FUNCTION_BLOCK FB_Startup
VAR_INPUT
END_VAR
VAR_OUTPUT
END_VAR
VAR
	timer1 : TON;
	timer2 : TON;
	timer3 : TON;
	timer4 : TON;
	timer5 : TON;
	timer6 : TON;
	timer7 : TON;
	EMG_STOP_RELEASED : BOOL;
END_VAR

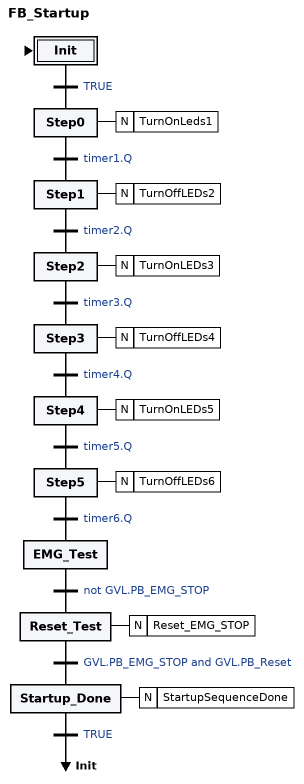
INITIAL_STEP Init:
END_STEP
TRANSITION FROM Init TO Step0
    := TRUE;
END_TRANSITION
STEP Step0:
    TurnOnLeds1(N);
END_STEP
TRANSITION FROM Step0 TO Step1
    := timer1.Q;
END_TRANSITION
STEP Step1:
    TurnOffLEDs2(N);
END_STEP
TRANSITION FROM Step1 TO Step2
    := timer2.Q;
END_TRANSITION
STEP Step2:
    TurnOnLEDs3(N);
END_STEP
TRANSITION FROM Step2 TO Step3
    := timer3.Q;
END_TRANSITION
STEP Step3:
    TurnOffLEDs4(N);
END_STEP
TRANSITION FROM Step3 TO Step4
    := timer4.Q;
END_TRANSITION
STEP Step4:
    TurnOnLEDs5(N);
END_STEP
TRANSITION FROM Step4 TO Step5
    := timer5.Q;
END_TRANSITION
STEP Step5:
    TurnOffLEDs6(N);
END_STEP
TRANSITION FROM Step5 TO EMG_Test
    := timer6.Q;
END_TRANSITION
STEP EMG_Test:
END_STEP
TRANSITION FROM EMG_Test TO Reset_Test
    := not GVL.PB_EMG_STOP;
END_TRANSITION
STEP Reset_Test:
    Reset_EMG_STOP(N);
END_STEP
TRANSITION FROM Reset_Test TO Startup_Done
    := GVL.PB_EMG_STOP and GVL.PB_Reset;
END_TRANSITION
STEP Startup_Done:
    StartupSequenceDone(N);
END_STEP
TRANSITION FROM Startup_Done TO Init
    := TRUE;
END_TRANSITION

METHOD AllLEDsTrigger : BOOL
VAR_INPUT
	OnOff : BOOL; // OnOff - Turn off, True - Turn On
END_VAR
GVL.LED_Comm_Fault := OnOff;
GVL.LED_EE_Grip := OnOff;
GVL.LED_EE_Ungrip := OnOff;
GVL.LED_EMG_STOP := OnOff;
GVL.LED_J1_CCW := OnOff;
GVL.LED_J1_CW := OnOff;
GVL.LED_J2_CCW := OnOff;
GVL.LED_J2_CW := OnOff;
GVL.LED_J3_CCW := OnOff;
GVL.LED_J3_CW := OnOff;
GVL.LED_Record_Delay := OnOff;
GVL.LED_Record_Pos := OnOff;
GVL.LED_Reset := OnOff;
GVL.LED_Start_Pause := OnOff;
GVL.LED_Warning := OnOff;
END_METHOD

ACTION Reset_EMG_STOP:
IF NOT GVL.PB_EMG_STOP THEN
	GVL.LED_EMG_STOP := TRUE;
END_IF

IF GVL.PB_EMG_STOP THEN
	GVL.LED_EMG_STOP := FALSE;
	GVL.LED_Reset := TRUE;
END_IF
END_ACTION

ACTION StartupSequenceDone:
GVL.LED_EMG_STOP := FALSE;
GVL.LED_Reset := FALSE;
GVL.system_state := state_enum.jog_joint_mode;
END_ACTION

ACTION TurnOffLEDs2:
timer1(IN := FALSE, PT := T#1S);
timer2(IN := TRUE, PT := T#1S);
timer3(IN := FALSE, PT := T#1S);
timer4(IN := FALSE, PT := T#1S);
timer5(IN := FALSE, PT := T#1S);
timer6(IN := FALSE, PT := T#1S);
timer7(IN := FALSE, PT := T#1S);
AllLEDsTrigger(FALSE);
END_ACTION

ACTION TurnOffLEDs4:
timer1(IN := FALSE, PT := T#1S);
timer2(IN := FALSE, PT := T#1S);
timer3(IN := FALSE, PT := T#1S);
timer4(IN := TRUE, PT := T#1S);
timer5(IN := FALSE, PT := T#1S);
timer6(IN := FALSE, PT := T#1S);
timer7(IN := FALSE, PT := T#1S);
AllLEDsTrigger(FALSE);
END_ACTION

ACTION TurnOffLEDs6:
timer1(IN := FALSE, PT := T#1S);
timer2(IN := FALSE, PT := T#1S);
timer3(IN := FALSE, PT := T#1S);
timer4(IN := FALSE, PT := T#1S);
timer5(IN := FALSE, PT := T#1S);
timer6(IN := TRUE, PT := T#1S);
timer7(IN := FALSE, PT := T#1S);
AllLEDsTrigger(FALSE);
END_ACTION

ACTION TurnOnLeds1:
timer1(IN := TRUE, PT := T#1S);
timer2(IN := FALSE, PT := T#1S);
timer3(IN := FALSE, PT := T#1S);
timer4(IN := FALSE, PT := T#1S);
timer5(IN := FALSE, PT := T#1S);
timer6(IN := FALSE, PT := T#1S);
timer7(IN := FALSE, PT := T#1S);
AllLEDsTrigger(TRUE);
END_ACTION

ACTION TurnOnLEDs3:
timer1(IN := FALSE, PT := T#1S);
timer2(IN := FALSE, PT := T#1S);
timer3(IN := TRUE, PT := T#1S);
timer4(IN := FALSE, PT := T#1S);
timer5(IN := FALSE, PT := T#1S);
timer6(IN := FALSE, PT := T#1S);
timer7(IN := FALSE, PT := T#1S);
AllLEDsTrigger(TRUE);
END_ACTION

ACTION TurnOnLEDs5:
timer1(IN := TRUE, PT := T#1S);
timer2(IN := FALSE, PT := T#1S);
timer3(IN := FALSE, PT := T#1S);
timer4(IN := FALSE, PT := T#1S);
timer5(IN := TRUE, PT := T#1S);
timer6(IN := FALSE, PT := T#1S);
timer7(IN := FALSE, PT := T#1S);
AllLEDsTrigger(TRUE);
END_ACTION

END_FUNCTION_BLOCK

(* stored: Version 1.1.0.1, ProductVersion 3.1.4024.13
   POU FB_Startup: Id {b471f5ac-fd76-4804-a6d3-9f17a23e0d1e}, SpecialFunc None
   Method AllLEDsTrigger: Id {56fddde5-8487-4a2d-a6eb-629934013dab}
   Action Reset_EMG_STOP: Id {e1a059ca-e1cc-40cf-b2b9-581c8d3cee73}
   Action StartupSequenceDone: Id {6d9cf29d-3216-46dd-8235-cc2d0bb2ba3d}
   Action TurnOffLEDs2: Id {001592bf-51e2-4ce1-8792-c625bfe1889c}
   Action TurnOffLEDs4: Id {f1f0bdb5-b6d0-4fba-80bf-214b3ce221e1}
   Action TurnOffLEDs6: Id {6d7c75b9-78c3-40d5-b315-14c6ad92b5f2}
   Action TurnOnLeds1: Id {9770b222-a122-43ae-9df8-13ef0f886ac4}
   Action TurnOnLEDs3: Id {fb04b18c-dfbf-4342-ab60-ff96bfa779fd}
   Action TurnOnLEDs5: Id {b4fc5097-dd0f-44dd-891c-f3cd7fb2d890} *)
